(* PLC project POC_ImportTest.xml, CODESYS CODESYS V3.5 SP19 Patch 1 *)
(* stored: creationDateTime 2026-07-04T00:00:00.0000000, modificationDateTime 2026-07-04T00:00:00.0000000 *)

(* ═══════════════════════════════════════════════════════════════ 🧪 ST_POC_ImportTest — Objet JETABLE, uniquement pour tester le mécanisme d'import PLCopenXML (GUID neuf, nom neuf, sans lien avec le programme réel). À supprimer du projet CODESYS après le test. Voir README.md du dossier test_import_poc/ pour le protocole d'observation. ═══════════════════════════════════════════════════════════════ *)
TYPE ST_POC_ImportTest : STRUCT
  Counter : INT := 0;  (* POC — compteur incrémenté à chaque appel avec Enable=TRUE *)
  Label : STRING(20);  (* POC — libellé texte, écrit par le FB de test *)
  Ready : BOOL;  (* POC — passe à TRUE après le premier appel réussi *)
END_STRUCT;
END_TYPE

(* ═══════════════════════════════════════════════════════════════ 🧪 FB_POC_ImportTest — Objet JETABLE, uniquement pour tester le mécanisme d'import PLCopenXML (GUID neuf, nom neuf, sans lien avec le programme réel). Ne pas appeler depuis un vrai programme métier. À supprimer du projet CODESYS après le test. Voir README.md du dossier test_import_poc/. ═══════════════════════════════════════════════════════════════ *)
FUNCTION_BLOCK FB_POC_ImportTest
  VAR_INPUT
    Enable : BOOL;  (* POC — active l'incrémentation du compteur *)
  END_VAR
  VAR_OUTPUT
    Done : BOOL;  (* POC — TRUE tant qu'Enable est actif *)
  END_VAR
  VAR_IN_OUT
    Data : ST_POC_ImportTest;  (* POC — structure de test lue/écrite par ce FB (VAR_IN_OUT) *)
  END_VAR

            
// 🧪 POC — logique volontairement minimale, sert juste à exercer le mécanisme d'import.
IF Enable THEN
    Data.Counter := Data.Counter + 1;
    Data.Label := 'POC_TEST';
    Data.Ready := TRUE;
    Done := TRUE;
ELSE
    Done := FALSE;
END_IF;

          
END_FUNCTION_BLOCK
